// TIA Portal V18 export
DATA_BLOCK "DB_Sensors"   // DB11
// stored: InstanceOfName FB_Sensors, InstanceOfType FB
"FB_Sensors"
   // VAR
   //    voltage_HL : Real;
   //    voltage_LL : Real;
   //    distance_HL : Real;
   //    distance_LL : Real;
   //    analogValue : Int;
   //    voltageOutput : Real;
   //    distanceOutput : Real;
   //    timeDelay : Time;
   //    "timer" : TP_TIME;
   //    trig : R_TRIG;
   //    startCond { S7_SetPoint := 'True'} : Bool;
   //    state : Bool;
   // END_VAR
BEGIN
END_DATA_BLOCK
